FUNCTION_BLOCK FB_DutyCycle
VAR_INPUT
	bEnable		: BOOL;
	fBaseTime	: REAL:=5.0; // [sec] min>0
	fOn_Duty	: REAL:=10.0; //min =0, max=100
END_VAR
VAR_OUTPUT
	bOut: BOOL;
END_VAR
VAR
	tBaseTime: TIME;
	ton_OnDuty: TON;
	fOnTime: REAL;
	tOnTime: TIME;
END_VAR


tBaseTime:=REAL_TO_TIME(fBaseTime*1000);
ton_OnDuty(PT:=tBaseTime,IN:=NOT ton_OnDuty.Q AND bEnable);

IF fOn_Duty<0 THEN;
	fOn_Duty:=0;
ELSIF fOn_Duty>100 THEN;
	fOn_Duty:=1000;
END_IF
	
fOnTime:=fBaseTime*fOn_Duty/100.0;
tOnTime:=REAL_TO_TIME(fOnTime*1000);

IF bEnable THEN;
	IF fOn_Duty<=0 THEN;
		bOut:=FALSE;
	ELSIF fOn_Duty>=100 THEN;
		bOut:=TRUE;
	ELSE;
		IF ton_OnDuty.ET<tOnTime THEN;
			bOut:=TRUE;
		ELSE
			bOut:=FALSE;
		END_IF		
	END_IF	
ELSE;
	bOut:=FALSE;
END_IF

END_FUNCTION_BLOCK

(* stored: Version 1.1.0.1, ProductVersion 3.1.4024.12
   POU FB_DutyCycle: Id {41274de3-ab3e-444e-8b5e-8fcc6e91c102}, SpecialFunc None *)
